// Mock of the dome (I_Dome): the commands only count, nothing moves.
FUNCTION_BLOCK FB_DomeMock IMPLEMENTS BROTLib.I_Dome
VAR
	bFailed		: BOOL;
	bIsParked	: BOOL := TRUE;
	bIsTracking	: BOOL;
	fPos		: LREAL;
	eShutter	: BROTLib.E_RoofState;
	nParkCalls	: UINT;
	nTrackCalls	: UINT;
END_VAR

METHOD Close : BOOL
Close := TRUE;
END_METHOD

METHOD Open : BOOL
Open := TRUE;
END_METHOD

METHOD Park : BOOL
nParkCalls := nParkCalls + 1;
bIsParked := TRUE;
bIsTracking := FALSE;
Park := TRUE;
END_METHOD

METHOD Reset : BOOL
bFailed := FALSE;
Reset := TRUE;
END_METHOD

METHOD Stop : BOOL
Stop := TRUE;
END_METHOD

METHOD StopTrack : BOOL
bIsTracking := FALSE;
StopTrack := TRUE;
END_METHOD

METHOD Track : BOOL
nTrackCalls := nTrackCalls + 1;
bIsParked := FALSE;
bIsTracking := TRUE;
Track := TRUE;
END_METHOD

PROPERTY Capabilities : INT
GET
Capabilities := 0;
END_GET
END_PROPERTY

PROPERTY Error : BOOL
GET
Error := bFailed;
END_GET
END_PROPERTY

PROPERTY ErrorID : UDINT
GET
ErrorID := 0;
END_GET
END_PROPERTY

PROPERTY Parked : BOOL
GET
Parked := bIsParked;
END_GET
END_PROPERTY

PROPERTY Position : LREAL
GET
Position := fPos;
END_GET
SET
fPos := Position;
END_SET
END_PROPERTY

PROPERTY RotState : BROTLib.E_DomeRotationState
GET
RotState := BROTLib.E_DomeRotationState.idle;
END_GET
END_PROPERTY

PROPERTY ShutterState : BROTLib.E_RoofState
GET
ShutterState := eShutter;
END_GET
SET
eShutter := ShutterState;
END_SET
END_PROPERTY

PROPERTY Tracking : BOOL
GET
Tracking := bIsTracking;
END_GET
END_PROPERTY

END_FUNCTION_BLOCK

(* stored: Version 1.1.0.1, ProductVersion 3.1.4024.15
   POU FB_DomeMock: Id {74b5e9c4-aee8-474a-82a8-2fd18e1b13fe}, SpecialFunc None
   Method Close: Id {2129f179-031c-4f16-bd66-db81fa9b1005}
   Method Open: Id {20583fa2-bb60-4421-a846-f8ae6a5b394d}
   Method Park: Id {612c7cbe-c374-40fc-aee3-0dd3942dd3aa}
   Method Reset: Id {07dd30a6-7dd2-47ae-bbb3-5c4ccb3770b5}
   Method Stop: Id {5177b14e-dec0-4c85-bd3d-17b5bcaca6c1}
   Method StopTrack: Id {f6d30648-cb35-4ad5-b22a-d2bb57129016}
   Method Track: Id {f8ee75c3-d379-4942-94af-1349be030839}
   Property Capabilities: Id {03a7f995-12ef-4a2c-b156-e33d3ea8554b}
   Get Get: Id {8e33c849-7617-492e-ae36-d0ede0ddb282}
   Property Error: Id {4f30c872-0f26-4bbf-b89c-0da617b5700b}
   Get Get: Id {d7f504c5-464f-4ef2-9a67-f4eb5c50992a}
   Property ErrorID: Id {ae8fbed9-2924-4324-a9dd-698112f6333d}
   Get Get: Id {202c93bd-bfa5-4566-9582-4063ab8d4e4a}
   Property Parked: Id {1d6f7c32-a789-4e79-9546-3a29a10b5397}
   Get Get: Id {18b6ee3c-221c-4155-97ff-83a4f1618aa8}
   Property Position: Id {224850c9-b26e-42a4-9a47-7d0c92bee7ff}
   Get Get: Id {b641347a-8ff8-445e-a2b6-dcee8fb3761a}
   Set Set: Id {b7b0b915-5512-4dca-bf2e-a75edf053aed}
   Property RotState: Id {1c9ce2fb-354e-47d0-8b14-4858c85f7387}
   Get Get: Id {164b626b-44f4-4a14-8d2a-602ac13d2afa}
   Property ShutterState: Id {fe66c2d3-1a0b-4cb6-a946-327c65b64388}
   Get Get: Id {2b0a14fe-3f82-4bce-8df3-40c70fb2665e}
   Set Set: Id {277f1e06-73aa-4701-8b4d-5b60b2264ac8}
   Property Tracking: Id {e46826cf-7133-4a7a-9ba5-ef975eb49554}
   Get Get: Id {4e56767f-2f6e-4f66-8b83-c7a9c0367dfe} *)
